ABB RAPID module: Count_only_pause.mod

%%%
  VERSION:1
  LANGUAGE:ENGLISH
%%%
MODULE MOD_Count_only_pause

    ! -------------------------------
    ! Define customized variables here
    ! ...

	! Tool variables:

	! Reference variables:

	PROC Main()
		ConfJ \On;
		ConfL \Off;
		! Program generated by RoboDK v6.0.7 for ABB IRB 120-3/0.6 on XX/XX/XXXX 12:58:43
		! Using nominal kinematics.
		WaitTime 0.100;
	ENDPROC

ENDMODULE
